Fanuc KAREL source: KA00106.KL

PROGRAM KA00106
%NOLOCKGROUP
VAR
  SRC: VECTOR
  DST: CONFIG
BEGIN
  SRC.X = 1.0
  DST = SRC
END KA00106
